FUNCTION_BLOCK FILL_CTRL (* Tank fill controller, written by hand *)
  (* Standard: 61499-2 *)
  (* Version 1.0, 2026-11-06, st2fb *)
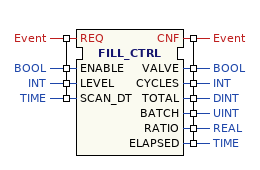
  EVENT_INPUT
    REQ WITH ENABLE, LEVEL, SCAN_DT;
  END_EVENT
  EVENT_OUTPUT
    CNF WITH VALVE, CYCLES, TOTAL, BATCH, RATIO, ELAPSED;
  END_EVENT
  VAR_INPUT
    ENABLE : BOOL;
    LEVEL : INT;
    SCAN_DT : TIME;
  END_VAR
  VAR_OUTPUT
    VALVE : BOOL;
    CYCLES : INT;
    TOTAL : DINT := 100;
    BATCH : UINT;
    RATIO : REAL;
    ELAPSED : TIME;
  END_VAR
  VAR
    LIMIT_LEVEL : INT := 10;
    I : INT;
  END_VAR
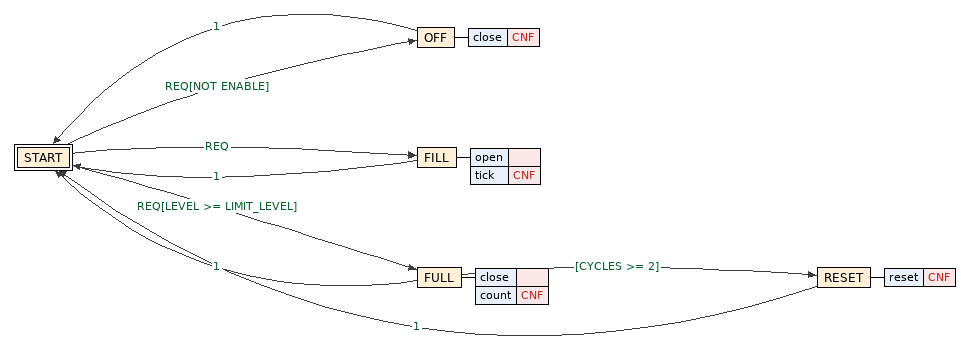
  EC_STATES
    START;
    OFF : close -> CNF;
    FILL : open, tick -> CNF;
    FULL : close, count -> CNF;
    RESET : reset -> CNF;
  END_STATES
  EC_TRANSITIONS
    START TO OFF := REQ[NOT ENABLE];
    START TO FULL := REQ[LEVEL >= LIMIT_LEVEL];
    START TO FILL := REQ;
    OFF TO START := 1;
    FILL TO START := 1;
    FULL TO RESET := [CYCLES >= 2];
    FULL TO START := 1;
    RESET TO START := 1;
  END_TRANSITIONS
  ALGORITHM close IN ST:
VALVE := FALSE;
  END_ALGORITHM
  ALGORITHM open IN ST:
VALVE := TRUE;
RATIO := RATIO + 0.5;
  END_ALGORITHM
  ALGORITHM tick IN ST:
ELAPSED := ELAPSED + SCAN_DT;
CASE LEVEL OF
  0: TOTAL := TOTAL + 1;
  1, 2: TOTAL := TOTAL + 10;
  3..5: TOTAL := TOTAL + 100;
  ELSE TOTAL := TOTAL - 1;
END_CASE;
  END_ALGORITHM
  ALGORITHM count IN ST:
CYCLES := CYCLES + 1;
FOR I := 1 TO 3 DO
  BATCH := BATCH + 2;
END_FOR;
WHILE BATCH > 4 DO
  BATCH := BATCH - 1;
END_WHILE;
  END_ALGORITHM
  ALGORITHM reset IN ST:
CYCLES := 0;
ELAPSED := T#0s;
  END_ALGORITHM
END_FUNCTION_BLOCK
